                //Check communication service: 0:UDP, 1:TCP, 2:LCOM
                IF (#diagnostics.localConfig.connection.comService = 16#01) THEN
                    //Communication service --> transport protocol TCP
                    #statTconPar.ConnectionType := 16#0B;
                    #diagnostics.localConfig.connection.useLComProtocol := FALSE;
                ELSIF (#diagnostics.localConfig.connection.comService = 16#02) THEN
                    //Communication service --> transport protocol TCP and LCom protocol
                    #statTconPar.ConnectionType := 16#0B;
                    #diagnostics.localConfig.connection.useLComProtocol := TRUE;
                ELSE
                    //Communication service --> NOT OK
                    //Write diagnostics
                    #statDiag.bufferIndex := #statDiag.bufferIndex + 1;
                    #statDiag.buffer[#statDiag.bufferIndex].status := ;
                    #statDiag.buffer[#statDiag.bufferIndex].subFunctionErrorID := 16#0000;
                    #statDiag.buffer[#statDiag.bufferIndex].additionalValue1 := #diagnostics.localConfig.connection.comService;//value from operator
                    #statDiag.buffer[#statDiag.bufferIndex].additionalValue2 := 0.0;
                    #statDiag.buffer[#statDiag.bufferIndex].additionalValue3 := 0.0;
                    #statDiag.buffer[#statDiag.bufferIndex].additionalValue4 := T#0ms;

                    #statState.connection := ;
                    GOTO ;
                END_IF;

                //Check unique connection identifier (16#0001...16#0FFF)
                IF ((#diagnostics.localConfig.connection.connectionID > 0)
                    AND
                    (#diagnostics.localConfig.connection.connectionID <= 4095))
                THEN
                    //Connection identifier -->OK
                    #statTconPar.ID := #diagnostics.localConfig.connection.connectionID;
                ELSE
                    //Connection identifier --> NOT OK
                    //Write diagnostics
                    #statDiag.bufferIndex := #statDiag.bufferIndex + 1;
                    #statDiag.buffer[#statDiag.bufferIndex].status := ;
                    #statDiag.buffer[#statDiag.bufferIndex].subFunctionErrorID := 16#0000;
                    #statDiag.buffer[#statDiag.bufferIndex].additionalValue1 := WORD_TO_UDINT(#diagnostics.localConfig.connection.connectionID);//value from user
                    #statDiag.buffer[#statDiag.bufferIndex].additionalValue2 := 0.0;
                    #statDiag.buffer[#statDiag.bufferIndex].additionalValue3 := 0.0;
                    #statDiag.buffer[#statDiag.bufferIndex].additionalValue4 := T#0ms;

                    #statState.connection := ;
                    GOTO ;
                END_IF;

                //check connection type: 1 = IPv4, 10 = QDN
                IF (#diagnostics.localConfig.connection.connectType = ) THEN
                    //connection type IPv4
                    ;
                ELSIF (#diagnostics.localConfig.connection.connectType = ) THEN
                    //connection type fully qualified domain name (QDN)
                    ;
                ELSE
                    //connection type --> NOT OK
                    //write diagnostics
                    #statDiag.bufferIndex := #statDiag.bufferIndex + 1;
                    #statDiag.buffer[#statDiag.bufferIndex].status := ;
                    #statDiag.buffer[#statDiag.bufferIndex].subFunctionErrorID := 16#0000;
                    #statDiag.buffer[#statDiag.bufferIndex].additionalValue1 := #diagnostics.localConfig.connection.connectType;//value from operator
                    #statDiag.buffer[#statDiag.bufferIndex].additionalValue2 := 0.0;
                    #statDiag.buffer[#statDiag.bufferIndex].additionalValue3 := 0.0;
                    #statDiag.buffer[#statDiag.bufferIndex].additionalValue4 := T#0ms;

                    #statState.connection := ;
                    GOTO ;
                END_IF;

                //If client
                IF (#diagnostics.localConfig.connection.isClient) THEN
                    //Partner port and remote address is not checked here
                    //The TCON will rise an error and return value, when the parameters (partnerPort or partnerIP) are wrong
                    //differ between different connection types (IPv4, QDN)
                    IF (#diagnostics.localConfig.connection.connectType = ) THEN
                        //remote addressing via IPv4
                        #statTconPar.RemotePort := #diagnostics.localConfig.connection.partnerPort;
                        #statTconPar.RemoteAddress := #diagnostics.localConfig.connection.partnerIP;
                    ELSE
                        //remote addressing via qualified domain name
                        #statTconParQdn.RemotePort := #diagnostics.localConfig.connection.partnerPort;
                        #statTconParQdn.RemoteQDN := #diagnostics.localConfig.connection.partnerQDN;
                        //additionally store all TCON configurations done before for QDN connection parameters
                        #statTconParQdn.ConnectionType := 16#0B;
                        #statTconParQdn.LocalPort := #diagnostics.localConfig.connection.localPort;
                        #statTconParQdn.InterfaceId := #diagnostics.localConfig.connection.interfaceID;
                        #statTconParQdn.ID := #diagnostics.localConfig.connection.connectionID;
                    END_IF;
                    //If server
                ELSE
                    //Accept requests from all partners or only specified partner is allowed
                    IF (#diagnostics.localConfig.connection.acceptUnknownPartner) THEN
                        //Accept requests from all partners
                        //differ between different connection types (IPv4, QDN)
                        IF (#diagnostics.localConfig.connection.connectType = ) THEN
                            #statTconPar.RemoteAddress.ADDR[1] := 0;
                            #statTconPar.RemoteAddress.ADDR[2] := 0;
                            #statTconPar.RemoteAddress.ADDR[3] := 0;
                            #statTconPar.RemoteAddress.ADDR[4] := 0;
                            #statTconPar.RemotePort := 0;
                        ELSE    //#CON_TYPE_QDN
                            #statTconParQdn.RemoteQDN := '';
                            #statTconParQdn.RemotePort := 0;
                        END_IF;
                    ELSE
                        //Only specified partner is allowed
                        //differ between different connection types (IPv4, QDN)
                        IF (#diagnostics.localConfig.connection.connectType = ) THEN
                            #statTconPar.RemoteAddress := #diagnostics.localConfig.connection.partnerIP;
                            #statTconPar.RemotePort := #diagnostics.localConfig.connection.partnerPort;
                        ELSE    //#CON_TYPE_QDN
                            #statTconParQdn.RemoteQDN := #diagnostics.localConfig.connection.partnerQDN;
                            #statTconParQdn.RemotePort := #diagnostics.localConfig.connection.partnerPort;
                        END_IF;
                    END_IF;
                END_IF;

                //Check cycleTime
                IF ((#diagnostics.localConfig.sender.cycleTime >= T#0ms)
                    AND
                    (#diagnostics.localConfig.sender.cycleTime <= T#+24d20h31m23s647ms))
                THEN
                    ;//CycleTime --> OK
                ELSE
                    //CycleTime --> NOT OK
                    #statDiag.bufferIndex := #statDiag.bufferIndex + 1;
                    #statDiag.buffer[#statDiag.bufferIndex].status := ;
                    #statDiag.buffer[#statDiag.bufferIndex].subFunctionErrorID := 16#0000;
                    #statDiag.buffer[#statDiag.bufferIndex].additionalValue1 := 0.0;
                    #statDiag.buffer[#statDiag.bufferIndex].additionalValue2 := 0.0;
                    #statDiag.buffer[#statDiag.bufferIndex].additionalValue3 := 0.0;
                    #statDiag.buffer[#statDiag.bufferIndex].additionalValue4 := #diagnostics.localConfig.sender.cycleTime;//value from operator

                    #statState.connection := ;
                    GOTO ;
                END_IF;

                //With LCom header
                IF (#diagnostics.localConfig.connection.useLComProtocol) THEN

                    //Check lifeSignCycleTime
                    IF ((#diagnostics.localConfig.connection.lifeSignCycleTime > T#0ms) //(1ms...T#+24d20h31m23s647ms)
                        AND
                        (#diagnostics.localConfig.connection.lifeSignCycleTime <= T#+24d20h31m23s647ms))
                    THEN
                        ;//lifeSignCycleTime--> OK
                    ELSE
                        //LifeSignCycle --> NOT OK
                        #statDiag.bufferIndex := #statDiag.bufferIndex + 1;
                        #statDiag.buffer[#statDiag.bufferIndex].status := ;
                        #statDiag.buffer[#statDiag.bufferIndex].subFunctionErrorID := 16#0000;
                        #statDiag.buffer[#statDiag.bufferIndex].additionalValue1 := 0.0;
                        #statDiag.buffer[#statDiag.bufferIndex].additionalValue2 := 0.0;
                        #statDiag.buffer[#statDiag.bufferIndex].additionalValue3 := 0.0;
                        #statDiag.buffer[#statDiag.bufferIndex].additionalValue4 := #diagnostics.localConfig.connection.lifeSignCycleTime;//value from operator

                        #statState.connection := ;
                        GOTO ;
                    END_IF;

                    //Check ackTimeOut
                    IF ((#diagnostics.localConfig.sender.ackTimeout > T#0ms)
                        AND
                        (#diagnostics.localConfig.sender.ackTimeout <= T#+24d20h31m23s647ms))
                    THEN
                        ;//AckTimeOut --> OK
                    ELSE
                        //AckTimeOut --> NOT OK
                        #statDiag.bufferIndex := #statDiag.bufferIndex + 1;
                        #statDiag.buffer[#statDiag.bufferIndex].status := ;
                        #statDiag.buffer[#statDiag.bufferIndex].subFunctionErrorID := 16#0000;
                        #statDiag.buffer[#statDiag.bufferIndex].additionalValue1 := 0.0;
                        #statDiag.buffer[#statDiag.bufferIndex].additionalValue2 := 0.0;
                        #statDiag.buffer[#statDiag.bufferIndex].additionalValue3 := 0.0;
                        #statDiag.buffer[#statDiag.bufferIndex].additionalValue4 := #diagnostics.localConfig.sender.ackTimeout;//value from operator

                        #statState.connection := ;
                        GOTO ;
                    END_IF;

                    //Check timeSync
                    IF (NOT #diagnostics.localConfig.timeSync.usePartnerTimestamps) THEN

                        IF ((#diagnostics.localConfig.timeSync.sendMode >= 0)//(0...2)
                            AND
                            (#diagnostics.localConfig.timeSync.sendMode <= 2))
                        THEN
                            CASE (#diagnostics.localConfig.timeSync.sendMode) OF

                                1: //TimeSync.cycleTime
                                    IF ((#diagnostics.localConfig.timeSync.cycleTime > T#0ms) //(1ms...T#+24d20h31m23s647ms)
                                        AND
                                        (#diagnostics.localConfig.timeSync.cycleTime <= T#+24d20h31m23s647ms))
                                    THEN
                                        ;//CycleTime --> OK
                                    ELSE
                                        //CycleTime --> Not OK
                                        #statDiag.bufferIndex := #statDiag.bufferIndex + 1;
                                        #statDiag.buffer[#statDiag.bufferIndex].status := ;
                                        #statDiag.buffer[#statDiag.bufferIndex].subFunctionErrorID := 16#0000;
                                        #statDiag.buffer[#statDiag.bufferIndex].additionalValue1 := 0.0;
                                        #statDiag.buffer[#statDiag.bufferIndex].additionalValue2 := 0.0;
                                        #statDiag.buffer[#statDiag.bufferIndex].additionalValue3 := 0.0;
                                        #statDiag.buffer[#statDiag.bufferIndex].additionalValue4 := #diagnostics.localConfig.timeSync.cycleTime;//value from user

                                        #statState.connection := ;
                                        GOTO ;

                                    END_IF;
                                2://TimeSync.sendAtTimeOfDay
                                    IF ((#diagnostics.localConfig.timeSync.sendAtTimeOfDay >= TOD#00:00:00.000) //(TOD#00:00:00.000...TOD#23:59:59.999)
                                        AND
                                        #diagnostics.localConfig.timeSync.sendAtTimeOfDay <= TOD#23:59:59.999)
                                    THEN
                                        ;//SendAtTimeOfDay --> OK
                                    ELSE
                                        //SendAtTimeOfDay --> NOT OK
                                        #statDiag.bufferIndex := #statDiag.bufferIndex + 1;
                                        #statDiag.buffer[#statDiag.bufferIndex].status := ;
                                        #statDiag.buffer[#statDiag.bufferIndex].subFunctionErrorID := 16#0000;
                                        #statDiag.buffer[#statDiag.bufferIndex].additionalValue1 := 0.0;
                                        #statDiag.buffer[#statDiag.bufferIndex].additionalValue2 := 0.0;
                                        #statDiag.buffer[#statDiag.bufferIndex].additionalValue3 := 0.0;
                                        #statDiag.buffer[#statDiag.bufferIndex].additionalValue4 := T#0ms;

                                        #statState.connection := ;
                                        GOTO ;
                                    END_IF;
                                ELSE
                                    ;
                            END_CASE;
                        ELSE
                            //SendMode --> NOT OK
                            #statDiag.bufferIndex := #statDiag.bufferIndex + 1;
                            #statDiag.buffer[#statDiag.bufferIndex].status := ;
                            #statDiag.buffer[#statDiag.bufferIndex].subFunctionErrorID := 16#0000;
                            #statDiag.buffer[#statDiag.bufferIndex].additionalValue1 := #diagnostics.localConfig.timeSync.sendMode;
                            #statDiag.buffer[#statDiag.bufferIndex].additionalValue2 := 0.0;
                            #statDiag.buffer[#statDiag.bufferIndex].additionalValue3 := 0.0;
                            #statDiag.buffer[#statDiag.bufferIndex].additionalValue4 := T#0ms;

                            #statState.connection := ;
                            GOTO ;
                        END_IF;
                    ELSE
                        //usePartnerTimeStamp

                        //Is sendMode inactive ?
                        IF #diagnostics.localConfig.timeSync.sendMode = 0 THEN
                            ;// Yes
                        ELSE
                            //SendMode --> NOT OK
                            #statDiag.bufferIndex := #statDiag.bufferIndex + 1;
                            #statDiag.buffer[#statDiag.bufferIndex].status := ;
                            #statDiag.buffer[#statDiag.bufferIndex].subFunctionErrorID := 16#0000;
                            #statDiag.buffer[#statDiag.bufferIndex].additionalValue1 := #diagnostics.localConfig.timeSync.sendMode;
                            #statDiag.buffer[#statDiag.bufferIndex].additionalValue2 := 0.0;
                            #statDiag.buffer[#statDiag.bufferIndex].additionalValue3 := 0.0;
                            #statDiag.buffer[#statDiag.bufferIndex].additionalValue4 := T#0ms;

                            #statState.connection := ;
                            GOTO ;
                        END_IF;

                    END_IF;
                ELSE
                    ;//No LCom Protocol is used
                END_IF;

                //differ between different connection types (IPv4, QDN)
                IF (#diagnostics.localConfig.connection.connectType = ) THEN
                    //IPv4
                    #instTCON(REQ := FALSE,
                              ID := #statTconPar.ID,
                              CONNECT := #statTconPar);
                    //store connection ID temporary
                    #tempConnOucId := #statTconPar.ID;
                ELSE
                    //QDN (CON_TYPE_QDN)
                    #instTCON(REQ := FALSE,
                              ID := #statTconParQdn.ID,
                              CONNECT := #statTconParQdn);
                    //store connection ID temporary
                    #tempConnOucId := #statTconParQdn.ID;
                END_IF;

                #instTSEND(REQ := FALSE,
                           ID := #tempConnOucId,
                           DATA := #statSend.tsendFct.data);

                #instTRCV(EN_R := FALSE,
                          ID := #tempConnOucId,
                          DATA := #statReceive.trcvFct.data);

                #instTDISCON(REQ := FALSE,
                             ID := #tempConnOucId);

                //Passive (server), active connection establishment (client)
                IF (#diagnostics.localConfig.connection.isClient) THEN
                    #statState.connection := ;
                    #statTconPar.ActiveEstablished := TRUE;
                    #statTconParQdn.ActiveEstablished := TRUE;
                ELSE
                    #statState.connection := ;
                    #statTconPar.ActiveEstablished := FALSE;
                    #statTconParQdn.ActiveEstablished := FALSE;
                END_IF;
            END_REGION INIT

        , :
            REGION OPEN_CLIENT_SERVER
                #instTCON.STATUS := 16#0000;

                //differ between different connection types (IPv4, QDN)
                IF (#diagnostics.localConfig.connection.connectType = ) THEN
                    //IPv4
                    #instTCON(REQ := TRUE,
                              CONNECT := #statTconPar,
                              ID := #diagnostics.localConfig.connection.connectionID);
                ELSE
                    //QDN (CON_TYPE_QDN)
                    #instTCON(REQ := TRUE,
                              CONNECT := #statTconParQdn,
                              ID := #diagnostics.localConfig.connection.connectionID);
                END_IF;

                // Error occurred
                IF (#instTCON.ERROR) THEN

                    //Local port is being used by the system
                    IF (#instTCON.STATUS = 16#80A2 OR (#diagnostics.localConfig.connection.connectType =  AND #statTconPar.LocalPort = 16#0)) THEN

                        #statDiag.bufferIndex := #statDiag.bufferIndex + 1;
                        #statDiag.buffer[#statDiag.bufferIndex].status := ;
                        #statDiag.buffer[#statDiag.bufferIndex].subFunctionErrorID := #instTCON.STATUS;
                        #statDiag.buffer[#statDiag.bufferIndex].additionalValue1 := #statTconPar.LocalPort;
                        #statDiag.buffer[#statDiag.bufferIndex].additionalValue2 := 0.0;
                        #statDiag.buffer[#statDiag.bufferIndex].additionalValue3 := 0.0;
                        #statDiag.buffer[#statDiag.bufferIndex].additionalValue4 := T#0ms;

                        #statState.connection := ;
                        GOTO ;
                        //Local port is being used by the system (in case of QDN)
                    ELSIF (#instTCON.STATUS = 16#80A2 OR (#diagnostics.localConfig.connection.connectType =  AND #statTconParQdn.LocalPort = 16#0)) THEN

                        #statDiag.bufferIndex := #statDiag.bufferIndex + 1;
                        #statDiag.buffer[#statDiag.bufferIndex].status := ;
                        #statDiag.buffer[#statDiag.bufferIndex].subFunctionErrorID := #instTCON.STATUS;
                        #statDiag.buffer[#statDiag.bufferIndex].additionalValue1 := #statTconParQdn.LocalPort;
                        #statDiag.buffer[#statDiag.bufferIndex].additionalValue2 := 0.0;
                        #statDiag.buffer[#statDiag.bufferIndex].additionalValue3 := 0.0;
                        #statDiag.buffer[#statDiag.bufferIndex].additionalValue4 := T#0ms;

                        #statState.connection := ;
                        GOTO ;
                    ELSIF (#instTCON.STATUS = 16#80B7 OR #instTCON.STATUS = 16#80A4) THEN
                        //IP address of the remote partner is invalid
                        #statDiag.bufferIndex := #statDiag.bufferIndex + 1;
                        #statDiag.buffer[#statDiag.bufferIndex].status := ;
                        #statDiag.buffer[#statDiag.bufferIndex].subFunctionErrorID := #instTCON.STATUS;
                        #statDiag.buffer[#statDiag.bufferIndex].additionalValue1 := 0.0;
                        #statDiag.buffer[#statDiag.bufferIndex].additionalValue2 := 0.0;
                        #statDiag.buffer[#statDiag.bufferIndex].additionalValue3 := 0.0;
                        #statDiag.buffer[#statDiag.bufferIndex].additionalValue4 := T#0ms;

                        #statState.connection := ;
                        GOTO ;
                    ELSIF (#instTCON.STATUS = 16#809B) THEN
                        //The local_device_id in the connection description does not match the CPU
                        #statDiag.bufferIndex := #statDiag.bufferIndex + 1;
                        #statDiag.buffer[#statDiag.bufferIndex].status := ;
                        #statDiag.buffer[#statDiag.bufferIndex].subFunctionErrorID := #instTCON.STATUS;
                        #statDiag.buffer[#statDiag.bufferIndex].additionalValue1 := UINT_TO_REAL(#diagnostics.localConfig.connection.interfaceID);//value from user
                        #statDiag.buffer[#statDiag.bufferIndex].additionalValue2 := 0.0;
                        #statDiag.buffer[#statDiag.bufferIndex].additionalValue3 := 0.0;
                        #statDiag.buffer[#statDiag.bufferIndex].additionalValue4 := T#0ms;

                        #statState.connection := ;
                        GOTO ;
                    ELSE
                        IF (#statState.connection = ) THEN

                            #statDiag.bufferIndex := #statDiag.bufferIndex + 1;
                            #statDiag.buffer[#statDiag.bufferIndex].status := ;
                            #statDiag.buffer[#statDiag.bufferIndex].subFunctionErrorID := #instTCON.STATUS;
                            #statDiag.buffer[#statDiag.bufferIndex].additionalValue1 := 0.0;
                            #statDiag.buffer[#statDiag.bufferIndex].additionalValue2 := 0.0;
                            #statDiag.buffer[#statDiag.bufferIndex].additionalValue3 := 0.0;
                            #statDiag.buffer[#statDiag.bufferIndex].additionalValue4 := T#0ms;

                            //Try reconnection after a wait time
                            #statIterator := 0;
                            #statState.connection := ;
                        ELSE
                            #statDiag.bufferIndex := #statDiag.bufferIndex + 1;
                            #statDiag.buffer[#statDiag.bufferIndex].status := ;
                            #statDiag.buffer[#statDiag.bufferIndex].subFunctionErrorID := #instTCON.STATUS;
                            //differ between different connection types (IPv4, QDN)
                            IF (#diagnostics.localConfig.connection.connectType = ) THEN
                                #statDiag.buffer[#statDiag.bufferIndex].additionalValue1 := #statTconPar.LocalPort;
                            ELSE    //CON_TYPE_QDN
                                #statDiag.buffer[#statDiag.bufferIndex].additionalValue1 := #statTconParQdn.LocalPort;
                            END_IF;
                            #statDiag.buffer[#statDiag.bufferIndex].additionalValue2 := 0.0;
                            #statDiag.buffer[#statDiag.bufferIndex].additionalValue3 := 0.0;
                            #statDiag.buffer[#statDiag.bufferIndex].additionalValue4 := T#0ms;

                            //Try reconnection after a wait time
                            #statIterator := 0;
                            #statState.connection := ;
                        END_IF;
                    END_IF;
                    //Job completed without error
                ELSIF (#instTCON.DONE) THEN

                    //Connection successfully established
                    #diagnostics.statistics.totalReconnects := #diagnostics.statistics.totalReconnects + 1;
                    #statState.connection := ;

                    #error := FALSE;

                    //Reset all state machines
                    #statState.receiver := ;
                    #statState.sender := ;
                    #statState.comReceiver := ;
                    #statState.comSender := ;
                    //Receive
                    #statReceive.trcvFct.dataOffset := 0;
                    #statReceive.trcvFct.dataLength := 0;
                    #statReceive.trcvFct.dataLengthRest := 0;
                    #statReceive.trcvFct.dataReceived := FALSE;
                    #statReceive.tempTelegram.index := 0;
                    #statReceive.tempTelegram.telegramType := 0;
                    #statReceive.numberOfLComHeader := 0;
                    #statReceive.dataTelegram.totalMessageLength := 0;
                    #statReceive.dataTelegram.actPackageLength := 0;
                    #statReceive.dataTelegram.ackMessageOffset := 0;
                    #statReceive.dataTelegram.messageOffset := 0;
                    #statReceive.dataTelegram.ackMessageCounter := 0;
                    #statReceive.dataTelegram.messageCounter := 0;
                    #statReceive.userData.totalLength := 0;
                    #statReceive.userData.offset := 0;
                    //Send
                    #statSend.tsendFct.dataLengthRest := 0;
                    #statSend.tsendFct.dataOffset := 0;
                    #statSend.tsendFct.status := 16#0000;
                    #statSend.expectedAck.package1.offset := 0;
                    #statSend.dataTelegram.messageCounter := 0;
                    #statSend.dataTelegram.ackMessageCounter := 0;
                    #statSend.dataTelegram.messageOffset := 0;
                    #statSend.dataTelegram.ackMessageOffset := 0;
                    #statSend.dataTelegram.actPackageLength := 0;
                    #statSend.dataTelegram.totalMessageLength := 0;
                    #statSend.numberOfLComPackage := 0;
                    #statSend.userData.totalLength := 0;
                    #statSend.userData.offset := 0;
                    #statSend.userData.sendCycleViolation := FALSE;
                    #statOldSend := FALSE;

                    #diagnostics.statistics.maxMsgSendingTime := T#0ms;
                    #diagnostics.localConfig.sender.cycleTime := T#0ms;
                    #diagnostics.localConfig.sender.ackTimeout := T#0ms;

                    #diagnostics.statistics.lastTimeSync.YEAR := 2200;
                    #statCopyNBytes := 0;

                    //Reset all timer
                    #instLocalLifeSignCycleTimer(IN := FALSE,
                                                 PT := #diagnostics.localConfig.connection.lifeSignCycleTime);

                    #instPartnerLifeSignCycleTimer(IN := FALSE,
                                                   PT := (#diagnostics.partnerConfig.connnection.lifeSignCycleTime));

                    #instLocalCycleTimeTimer(IN := FALSE,
                                             PT := #diagnostics.localConfig.sender.cycleTime);

                    #instExpectedAckPackage1(IN := FALSE,
                                             PT := #diagnostics.localConfig.sender.ackTimeout);

                    #instSyncTimer(IN := FALSE,
                                   PT := T#1s);

                    #instSendErrorTimer(IN := FALSE,
                                        PT := );

                    #instRcvErrorTimer(IN := FALSE,
                                       PT := );

                    //Reset all active failures in the diagnostics buffer
                    FOR #statIterator := 0 TO  BY 1 DO
                        #diagnostics.buffer[#statIterator].isActive := FALSE;
                    END_FOR;

                    //With LCom protocol
                    IF (#diagnostics.localConfig.connection.useLComProtocol = TRUE) THEN

                        IF (#statConnectAttempts MOD 2 = 0) THEN
                            //1st try LCom Version 2.0
                            #statActualLocalLComVersion := ;
                            #statSend.configTelegramV2.LComVersion := ;
                            #statSend.configTelegramV2.status := BOOL_TO_BYTE(#diagnostics.localConfig.timeSync.usePartnerTimestamps);
                            #statSend.configTelegramV2.sendModeSyncTime := #diagnostics.localConfig.timeSync.sendMode;
                            #statSend.configTelegramV2.lifeSignCycle := #diagnostics.localConfig.connection.lifeSignCycleTime;
                            #statSend.configTelegramV2.cycleTime := #configuration.sender.cycleTime;
                            #statSend.configTelegramV2.ackTimeOut := #configuration.sender.ackTimeout;
                            #statSend.configTelegramV2.maxSendDataLength := #diagnostics.localConfig.sizeOfSendBuffer;
                            #statSend.configTelegramV2.maxReceiveDataLength := #diagnostics.localConfig.sizeOfReceiveBuffer;

                            #statSend.dataTelegram.LComVersion := #statSend.configTelegramV2.LComVersion;
                        ELSE
                            //2nd try LCom Version 1.0
                            #statActualLocalLComVersion := ;
                            #statSend.configTelegramV1.LComVersion := ;
                            #statSend.configTelegramV1.comMode := 16#03;
                            #statSend.configTelegramV1.slidingWindow := 1;
                            #statSend.configTelegramV1.status := BOOL_TO_BYTE(#diagnostics.localConfig.timeSync.usePartnerTimestamps);
                            #statSend.configTelegramV1.sendModeSyncTime := #diagnostics.localConfig.timeSync.sendMode;

                            #statSend.dataTelegram.LComVersion := #statSend.configTelegramV1.LComVersion;

                            //Check max. lifeSignCycleTime
                            IF (#diagnostics.localConfig.connection.lifeSignCycleTime > T#65535ms) THEN

                                #statDiag.bufferIndex := #statDiag.bufferIndex + 1;
                                #statDiag.buffer[#statDiag.bufferIndex].additionalValue4 := #diagnostics.localConfig.connection.lifeSignCycleTime;
                                #diagnostics.localConfig.connection.lifeSignCycleTime := T#65535ms;

                                #statDiag.buffer[#statDiag.bufferIndex].status := ;
                                #statDiag.buffer[#statDiag.bufferIndex].subFunctionErrorID := 16#0000;
                                #statDiag.buffer[#statDiag.bufferIndex].additionalValue1 := 65535.0;
                                #statDiag.buffer[#statDiag.bufferIndex].additionalValue2 := 0.0;
                                #statDiag.buffer[#statDiag.bufferIndex].additionalValue3 := 0.0;
                            ELSE
                                ;
                            END_IF;
                            #statSend.configTelegramV1.lifeSignCycle := TIME_TO_UINT(#diagnostics.localConfig.connection.lifeSignCycleTime);

                            //Check max.sizeOfSendBuffer
                            IF (#diagnostics.localConfig.sizeOfSendBuffer > 65535) THEN
                                #diagnostics.localConfig.sizeOfSendBuffer := 65535;
                                #statSend.configTelegramV1.maxSendDataLength := 65535;
                            ELSE
                                #statSend.configTelegramV1.maxSendDataLength := UDINT_TO_UINT(#diagnostics.localConfig.sizeOfSendBuffer);
                            END_IF;

                            //Check max.sizeOfReceiveBuffer
                            IF (#diagnostics.localConfig.sizeOfReceiveBuffer > 65535) THEN
                                #diagnostics.localConfig.sizeOfReceiveBuffer := 65535;
                                #statSend.configTelegramV1.maxReceiveDataLength := 65535;
                            ELSE
                                #statSend.configTelegramV1.maxReceiveDataLength := UDINT_TO_UINT(#diagnostics.localConfig.sizeOfReceiveBuffer);
                            END_IF;

                        END_IF;
                        //Set telegram type of data telegrams for LCom Version 1.0 and 2.0
                        #statSend.dataTelegram.telegramType := 16#0A;

                        //Start sender config directly with LCom protocol
                        #statState.cfgSender := ;
                    ELSE
                        //without LCom
                        #statCompare.sender.cycleTime := #configuration.sender.cycleTime;
                        #diagnostics.localConfig.sender.cycleTime := #configuration.sender.cycleTime;

                        #diagnostics.partnerConfig.sizeOfReceiveBuffer := 0;
                        #diagnostics.partnerConfig.sizeOfSendBuffer := 0;
                        #connected := #statConnected := TRUE;
                        #statState.cfgSender := ;

                        #statDiag.bufferIndex := #statDiag.bufferIndex + 1;
                        #statDiag.buffer[#statDiag.bufferIndex].status := ;
                        #statDiag.buffer[#statDiag.bufferIndex].subFunctionErrorID := 16#0000;
                        #statDiag.buffer[#statDiag.bufferIndex].additionalValue1 := 0.0;
                        #statDiag.buffer[#statDiag.bufferIndex].additionalValue2 := 0.0;
                        #statDiag.buffer[#statDiag.bufferIndex].additionalValue3 := 0.0;
                        #statDiag.buffer[#statDiag.bufferIndex].additionalValue4 := T#0ms;
                    END_IF;
                    //TCON still in progress
                ELSE
                    IF (#diagnostics.localConfig.connection.isClient) THEN

                        #statDiag.bufferIndex := #statDiag.bufferIndex + 1;
                        #statDiag.buffer[#statDiag.bufferIndex].status := ;
                        #statDiag.buffer[#statDiag.bufferIndex].subFunctionErrorID := 16#0000;
                        #statDiag.buffer[#statDiag.bufferIndex].additionalValue1 := 0.0;
                        #statDiag.buffer[#statDiag.bufferIndex].additionalValue2 := 0.0;
                        #statDiag.buffer[#statDiag.bufferIndex].additionalValue3 := 0.0;
                        #statDiag.buffer[#statDiag.bufferIndex].additionalValue4 := T#0ms;
                    ELSE
                        #statDiag.bufferIndex := #statDiag.bufferIndex + 1;
                        #statDiag.buffer[#statDiag.bufferIndex].status := ;
                        #statDiag.buffer[#statDiag.bufferIndex].subFunctionErrorID := 16#0000;
                        #statDiag.buffer[#statDiag.bufferIndex].additionalValue1 := 0.0;
                        #statDiag.buffer[#statDiag.bufferIndex].additionalValue2 := 0.0;
                        #statDiag.buffer[#statDiag.bufferIndex].additionalValue3 := 0.0;
                        #statDiag.buffer[#statDiag.bufferIndex].additionalValue4 := T#0ms;
                    END_IF;
                END_IF;
            END_REGION OPEN_CLIENT_SERVER

        :
            REGION WAIT
                //Wait and then establish the connection
                IF (#statIterator > ) THEN

                    #tempConnOucId := 0;

                    //differ between different connection types (IPv4, QDN)
                    IF (#diagnostics.localConfig.connection.connectType = ) THEN
                        //IPv4
                        #instTCON(REQ := FALSE,
                                  ID := #statTconPar.ID,
                                  CONNECT := #statTconPar);
                        //store connection ID temporary
                        #tempConnOucId := #statTconPar.ID;
                    ELSE
                        //QDN (CON_TYPE_QDN)
                        #instTCON(REQ := FALSE,
                                  ID := #statTconParQdn.ID,
                                  CONNECT := #statTconParQdn);
                        //store connection ID temporary
                        #tempConnOucId := #statTconParQdn.ID;
                    END_IF;

                    #instTSEND(REQ := FALSE,
                               ID := #tempConnOucId,
                               DATA := #statSend.tsendFct.data);

                    #instTRCV(EN_R := FALSE,
                              ID := #tempConnOucId,
                              DATA := #statReceive.trcvFct.data);

                    #instTDISCON(REQ := FALSE,
                                 ID := #tempConnOucId);

                    IF (#diagnostics.localConfig.connection.isClient) THEN
                        #statState.connection := ;
                        #statTconPar.ActiveEstablished := TRUE;
                        #statTconParQdn.ActiveEstablished := TRUE;
                    ELSE
                        #statState.connection := ;
                        #statTconPar.ActiveEstablished := FALSE;
                        #statTconParQdn.ActiveEstablished := FALSE;
                    END_IF;

                ELSE
                    #statIterator := #statIterator + 1;
                END_IF;
            END_REGION WAIT

        :
            REGION FINISH_TSEND
                IF (#statIterator > ) THEN
                    #statIterator := 0;
                    #statState.connection := ;
                ELSE
                    //differ between different connection types (IPv4, QDN)
                    IF (#diagnostics.localConfig.connection.connectType = ) THEN
                        #tempConnOucId := #statTconPar.ID;
                    ELSE    //CON_TYPE_QDN
                        #tempConnOucId := #statTconParQdn.ID;
                    END_IF;

                    #instTSEND(REQ := TRUE,
                               LEN := #statSend.tsendFct.dataOffset,
                               ID := #tempConnOucId,
                               DATA := #statSend.tsendFct.data,
                               STATUS => #statSend.tsendFct.status);

                    IF ((#statSend.tsendFct.status = 16#0000) OR (#instTSEND.ERROR)) THEN
                        //"TSEND" instruction is finished
                        #statState.connection := ;
                    ELSE
                        ;//"TSEND" instruction still in process
                    END_IF;
                END_IF;
                #statIterator := #statIterator + 1;
            END_REGION FINISH_TSEND

        :
            REGION FINISH_TRCV

                IF (#statIterator > ) THEN
                    #statState.connection := ;
                ELSE
                    //differ between different connection types (IPv4, QDN)
                    IF (#diagnostics.localConfig.connection.connectType = ) THEN
                        #tempConnOucId := #statTconPar.ID;
                    ELSE    //CON_TYPE_QDN
                        #tempConnOucId := #statTconParQdn.ID;
                    END_IF;

                    #instTRCV(EN_R := TRUE,
                              ID := #tempConnOucId,
                              LEN := 0,
                              ADHOC := TRUE,
                              NDR => #statReceive.trcvFct.dataReceived,
                              RCVD_LEN => #statReceive.trcvFct.dataLength,
                              DATA := #statReceive.trcvFct.data);

                    //Is the "TRCV" instruction still in process
                    IF (#instTRCV.ERROR OR NOT #instTRCV.BUSY) THEN
                        #statState.connection := ;
                    ELSE
                        ;//TRCV instruction still in process
                    END_IF;
                END_IF;
                #statIterator := #statIterator + 1;
            END_REGION FINISH_TRCV

        :
            REGION CLOSE_CONNECTION
                //reset FB Outputs
                #connected := #statConnected := FALSE;
                #sending := #statSending := FALSE;
                #receivedDataLength := 0;
                #error := FALSE;

                //Is "TSEND" instruction still in process ?
                IF (#statSend.tsendFct.status <> 16#0000) THEN
                    //"TSEND" instruction still in process
                    #statState.connection := ;
                    #statIterator := 0;
                ELSE
                    ;//"TSEND" instruction is finished
                END_IF;

                #instTRCV(EN_R := TRUE,
                          ID := #diagnostics.localConfig.connection.connectionID,
                          LEN := 0,
                          ADHOC := TRUE,
                          NDR => #statReceive.trcvFct.dataReceived,
                          RCVD_LEN => #statReceive.trcvFct.dataLength,
                          DATA := #statReceive.trcvFct.data);

                //Is the "TRCV" instruction still in process
                IF (#instTRCV.ERROR OR NOT #instTRCV.BUSY) THEN
                    #statState.connection := ;
                ELSE
                    #statState.connection := ;
                    #statIterator := 0;
                END_IF;
            END_REGION CLOSE_CONNECTION

        :
            REGION CALL_TDISCON
                //differ between different connection types (IPv4, QDN)
                IF (#diagnostics.localConfig.connection.connectType = ) THEN
                    #tempConnOucId := #statTconPar.ID;
                ELSE    //CON_TYPE_QDN
                    #tempConnOucId := #statTconParQdn.ID;
                END_IF;

                #instTSEND(REQ := FALSE,
                           LEN := #statSend.tsendFct.dataOffset,
                           ID := #tempConnOucId,
                           DATA := #statSend.tsendFct.data);

                #instTRCV(EN_R := FALSE,
                          ID := #diagnostics.localConfig.connection.connectionID,
                          LEN := 0,
                          ADHOC := TRUE,
                          NDR => #statReceive.trcvFct.dataReceived,
                          RCVD_LEN => #statReceive.trcvFct.dataLength,
                          DATA := #statReceive.trcvFct.data);

                #instTDISCON(REQ := TRUE,
                             ID := #tempConnOucId);

                //Error occurred during processing
                IF (#instTDISCON.ERROR) THEN

                    #statDiag.bufferIndex := #statDiag.bufferIndex + 1;
                    #statDiag.buffer[#statDiag.bufferIndex].status := ;
                    #statDiag.buffer[#statDiag.bufferIndex].subFunctionErrorID := #instTDISCON.STATUS;
                    #statDiag.buffer[#statDiag.bufferIndex].additionalValue1 := 0.0;
                    #statDiag.buffer[#statDiag.bufferIndex].additionalValue2 := 0.0;
                    #statDiag.buffer[#statDiag.bufferIndex].additionalValue3 := 0.0;
                    #statDiag.buffer[#statDiag.bufferIndex].additionalValue4 := T#0ms;

                    #statState.connection := ;

                    #instTDISCON(REQ := FALSE,
                                 ID := #tempConnOucId);

                ELSIF (#instTDISCON.DONE) THEN

                    #instTDISCON(REQ := FALSE,
                                 ID := #tempConnOucId);
                    //Job executed without errors
                    IF (#enable AND (NOT #statFallingEdgeEnable)) THEN
                        //Reconnect automatically if not in disconnecting process
                        #statIterator := 0;
                        #statState.connection := ;
                    ELSE
                        //Reset all active failures in the diagnostics buffer
                        FOR #statIterator := 0 TO  BY 1 DO
                            #diagnostics.buffer[#statIterator].isActive := FALSE;
                        END_FOR;

                        #statState.connection := ;
                    END_IF;
                    //Job is not completed yet
                ELSE
                    ;//Wait until job is finished
                END_IF;
            END_REGION CALL_TDISCON

        :
            REGION ERROR
                ;
            END_REGION ERROR
    END_CASE;
END_REGION STATE_MACHINE

REGION DIAGNOSTICS
    // -----------------------------------------------------------------------------------------------------------
    //Diagnostics buffer
    // -----------------------------------------------------------------------------------------------------------
:
    //Diagnostics entry is in the temp. buffer
    IF (#statDiag.bufferIndex <> -1) THEN

        //Get current time
        #statRet := RD_LOC_T(#tempActTime);
        //init
        #statDiag.actualIndex := 0;

        WHILE (#statDiag.actualIndex <= #statDiag.bufferIndex) DO

            #tempUDint := 0;
            //Check if the failure is already in the buffer and still active
            FOR #statIterator := 0 TO  BY 1 DO

                IF (#diagnostics.buffer[#statIterator].isActive = TRUE) THEN

                    IF ((#statDiag.buffer[#statDiag.actualIndex].status = )
                        AND
                        (#diagnostics.buffer[#statIterator].status = )
                        AND
                        (#diagnostics.buffer[#statIterator].additionalValue1 = #statDiag.buffer[#statDiag.actualIndex].additionalValue1)
                        AND
                        (#diagnostics.buffer[#statIterator].additionalValue2 = #statDiag.buffer[#statDiag.actualIndex].additionalValue2)
                        AND
                        (#diagnostics.buffer[#statIterator].additionalValue3 = #statDiag.buffer[#statDiag.actualIndex].additionalValue3)) THEN
                        //Retrigger just the activation time
                        #diagnostics.buffer[#statIterator].timestamp := #tempActTime;
                        #diagnostics.buffer[#statIterator].additionalValue4 := #statDiag.buffer[#statDiag.actualIndex].additionalValue4;
                        #tempUDint := 100;
                        EXIT;
                    ELSIF ((#diagnostics.buffer[#statIterator].status = #statDiag.buffer[#statDiag.actualIndex].status)
                        AND
                        (#diagnostics.buffer[#statIterator].additionalValue1 = #statDiag.buffer[#statDiag.actualIndex].additionalValue1)
                        AND
                        (#diagnostics.buffer[#statIterator].additionalValue2 = #statDiag.buffer[#statDiag.actualIndex].additionalValue2)
                        AND
                        (#diagnostics.buffer[#statIterator].additionalValue3 = #statDiag.buffer[#statDiag.actualIndex].additionalValue3)
                        AND
                        (#diagnostics.buffer[#statIterator].additionalValue4 = #statDiag.buffer[#statDiag.actualIndex].additionalValue4)) THEN
                        //Retrigger just the activation time
                        #diagnostics.buffer[#statIterator].timestamp := #tempActTime;
                        #tempUDint := 100;
                        EXIT;
                    ELSE
                        ;//ErrorId is not in the diagnostics buffer
                    END_IF;
                END_IF;
            END_FOR;

            IF (#tempUDint = 100) THEN
                ;//ErrorId was already retriggered
            ELSE
                //Check range of diagnostics ring buffer [0...DIAG_ARRAY]
                IF ((#diagnostics.bufferIndex = 255) OR (#diagnostics.bufferIndex = )) THEN
                    #diagnostics.bufferIndex := 0;
                ELSE
                    #diagnostics.bufferIndex := #diagnostics.bufferIndex + 1;
                END_IF;

                //Stored new entry in the diagnostics buffer
                #diagnostics.buffer[#diagnostics.bufferIndex].status := #statDiag.buffer[#statDiag.actualIndex].status;
                #diagnostics.buffer[#diagnostics.bufferIndex].timestamp := #tempActTime;
                #diagnostics.buffer[#diagnostics.bufferIndex].isActive := TRUE;

                #diagnostics.buffer[#diagnostics.bufferIndex].subFunctionErrorID := #statDiag.buffer[#statDiag.actualIndex].subFunctionErrorID;
                #diagnostics.buffer[#diagnostics.bufferIndex].additionalValue1 := #statDiag.buffer[#statDiag.actualIndex].additionalValue1;
                #diagnostics.buffer[#diagnostics.bufferIndex].additionalValue2 := #statDiag.buffer[#statDiag.actualIndex].additionalValue2;
                #diagnostics.buffer[#diagnostics.bufferIndex].additionalValue3 := #statDiag.buffer[#statDiag.actualIndex].additionalValue3;
                #diagnostics.buffer[#diagnostics.bufferIndex].additionalValue4 := #statDiag.buffer[#statDiag.actualIndex].additionalValue4;
            END_IF;

            IF ((#diagnostics.buffer[#diagnostics.bufferIndex].status = )
                OR (#diagnostics.buffer[#diagnostics.bufferIndex].status = )
                OR (#diagnostics.buffer[#diagnostics.bufferIndex].status = ))
            THEN
                #statConnectAttempts := 0;
                #diagnostics.statistics.lastConnect := #tempActTime;
            END_IF;

            //Set FB status
            #status := #statStatus := #statDiag.buffer[#statDiag.actualIndex].status;

            //Check if FB.error has been set ?
            IF ((#statDiag.buffer[#statDiag.actualIndex].status >= )//16#8200
                AND
                (#statDiag.buffer[#statDiag.actualIndex].status <= ))//16#8614
            THEN

                #error := TRUE;
                #connected := #statConnected := FALSE;
                #sending := #statSending := FALSE;
                #dataReceived := #statDataReceived := FALSE;
                #receivedDataLength := 0;

                //Check if FB.busy has been set ?
                IF ((#statDiag.buffer[#statDiag.actualIndex].status >= )//16#8600
                    AND
                    (#statDiag.buffer[#statDiag.actualIndex].status <= ))//16#8614
                THEN
                    #busy := TRUE;
                ELSE
                    #busy := FALSE;
                END_IF;

                EXIT;//Leave loop
            ELSE
                ;
            END_IF;

            //Increase index
            #statDiag.actualIndex := #statDiag.actualIndex + 1;

        END_WHILE;
    ELSE
        ;//No failure
    END_IF;//End: Diagnostics buffer
END_REGION DIAGNOSTICS
END_FUNCTION_BLOCK